Staubli VAL3: utData.dtx

public num nVal
public bool bStatus
public string sSourceImg1
public string sSourceImg2
